Fanuc KAREL source: kd00068.KL

-- PROVISIONAL review KL for V1013-1; original PC SHA256 bce0d8b3e73cf6692d564c39646a4f04ab738961b3d16c2260da6a311af2ec7f
-- Incomplete behavior may be omitted. Consult companion uncertainty JSON. Do not deploy.
PROGRAM KD00068
%NOLOCKGROUP
VAR
  I : INTEGER
  J : INTEGER
  B : BOOLEAN
  R : REAL
  S : STRING[80]
BEGIN
  -- UNRESOLVED_PC offsets 5-29; opcodes 9D,81,18,9D,1B,9D,12,2E,1B,2E,13,04
  -- UNRESOLVED_PC offsets 34-38; opcodes 7F
END KD00068
